Fanuc KAREL source: kt00605.compact.KL

PROGRAM KT00605
%STACKSIZE=65535
%PRIORITY=65535
%NOLOCKGROUP
VAR
I1 : INTEGER
I2 : INTEGER
OUT : REAL
BEGIN
I1=2
I2=3
I1=2
I2=3
OUT=((-I1))
END KT00605
